Fanuc KAREL source: NC0062.KL

PROGRAM NC0062
%NOLOCKGROUP
ROUTINE R
VAR
S1:INTEGER;S2:INTEGER
BEGIN
--
S1=1
FOR S2=1 TO 2 DO
S1=(S1+1)
ENDFOR
END R
BEGIN
R
END NC0062
